Staubli VAL3: initText.pgx

public program initText(utText& x_utText, string x_sPage, string x_sId, string x_sType)
begin
  x_utText.Common.sPage=x_sPage
  x_utText.Common.sID=x_sId
  switch x_sType
    case "Num"
      userPageBind(x_utText.Common.sPage,x_utText.Common.sID,"value",x_utText.Common.nValue,1,"rw")
    break
    case "String"
      userPageBind(x_utText.Common.sPage,x_utText.Common.sID,"value",x_utText.Common.sValue,1,"rw")
    break
  endSwitch
  userPageBind(x_utText.Common.sPage,x_utText.Common.sID,"style.backgroundColor",x_utText.Appearance.sBackgroundColour,1,"r")
  //
  x_utText.Appearance.sBackgroundColour="trasparent"
  //
end
